FUNCTION_BLOCK ControlPanel (* Composite Function Block Type *)
  (* Standard: 61499-2 *)
  (* Version 0.0, 7/2/2026, template *)
  PACKAGE Main;
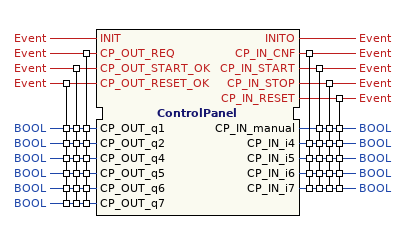
  EVENT_INPUT
    INIT; (* Initialization Request *)
    CP_OUT_REQ WITH CP_OUT_q1, CP_OUT_q2, CP_OUT_q4, CP_OUT_q5, CP_OUT_q6, CP_OUT_q7; (* Normal Execution Request *)
    CP_OUT_START_OK WITH CP_OUT_q1, CP_OUT_q2, CP_OUT_q4, CP_OUT_q5, CP_OUT_q6, CP_OUT_q7;
    CP_OUT_RESET_OK WITH CP_OUT_q1, CP_OUT_q2, CP_OUT_q4, CP_OUT_q5, CP_OUT_q6, CP_OUT_q7;
  END_EVENT
  EVENT_OUTPUT
    INITO; (* Initialization Confirm *)
    CP_IN_CNF WITH CP_IN_i4, CP_IN_i5, CP_IN_i6, CP_IN_i7; (* Execution Confirmation *)
    CP_IN_START WITH CP_IN_manual, CP_IN_i4, CP_IN_i5, CP_IN_i6, CP_IN_i7;
    CP_IN_STOP WITH CP_IN_manual, CP_IN_i4, CP_IN_i5, CP_IN_i6, CP_IN_i7;
    CP_IN_RESET WITH CP_IN_manual, CP_IN_i4, CP_IN_i5, CP_IN_i6, CP_IN_i7;
  END_EVENT
  VAR_INPUT
    CP_OUT_q1 : BOOL; (* Input event qualifier *)
    CP_OUT_q2 : BOOL;
    CP_OUT_q4 : BOOL;
    CP_OUT_q5 : BOOL;
    CP_OUT_q6 : BOOL;
    CP_OUT_q7 : BOOL;
  END_VAR
  VAR_OUTPUT
    CP_IN_manual : BOOL; (* Output event qualifier *)
    CP_IN_i4 : BOOL;
    CP_IN_i5 : BOOL;
    CP_IN_i6 : BOOL;
    CP_IN_i7 : BOOL;
  END_VAR
  FBS
    CP_OUT : ControlPanelOut;
    CP_IN : ControlPanelIn;
  END_FBS
  EVENT_CONNECTIONS
    INIT TO CP_OUT.CCD65B7F67E00C87;
    CP_OUT_REQ TO CP_OUT.4778653D8DBF7248;
    CP_OUT_START_OK TO CP_OUT.DC4AC429D7DC72F4;
    CP_OUT_RESET_OK TO CP_OUT.ADC8D44EE6F5CFC7;
    CP_OUT.F7D5ED5A0E4491B7 TO CP_IN.8DC0B17FED05A165;
    CP_IN.01AE14A4F2450C6A TO INITO;
    CP_IN.E44B3C7CBCF63ADC TO CP_IN_CNF;
    CP_IN.FE8C6726676F44CD TO CP_IN_START;
    CP_IN.D7A4A0CA0112ED64 TO CP_IN_STOP;
    CP_IN.2403870DB0D5CE05 TO CP_IN_RESET;
  END_CONNECTIONS
  DATA_CONNECTIONS
    CP_OUT_q1 TO CP_OUT.C26EC91ADA4C3749;
    CP_OUT_q2 TO CP_OUT.8B5737DEFF5224B0;
    CP_OUT_q4 TO CP_OUT.E98BCB8EC09F669C;
    CP_OUT_q5 TO CP_OUT.972C67A1D7FE12B3;
    CP_OUT_q6 TO CP_OUT.15CA038062847536;
    CP_OUT_q7 TO CP_OUT.BCF57BAEFF0C3E81;
    CP_IN.5C09E78C1FA53551 TO CP_IN_manual;
    CP_IN.EC38A52344DEA219 TO CP_IN_i4;
    CP_IN.B26F11C5711BF1BD TO CP_IN_i5;
    CP_IN.8C1851B751A1950C TO CP_IN_i6;
    CP_IN.0EEA07D7271FFC63 TO CP_IN_i7;
  END_CONNECTIONS
END_FUNCTION_BLOCK
